// TIA Portal V20 export
DATA_BLOCK "DB020_Com LabView"   // DB20
{ S7_Optimized_Access := 'FALSE' }
// stored: AutoNumber false
   VAR
      E_Lebenszeichen : DInt := 0;   // E_Lebenszeichen
      E_Rückmeldung_Startfreigabe_Zwischenbefundung_erhalten : Bool;   // E_Rückmeldung_Startfreigabe_Zwischenbefundung_erhalten
      E_Rückmeldung_Zwischenbefundung_fertig : Bool;   // E_Rückmeldung_Zwischenbefundung_fertig
      "E_Messgerät ist bereit und verbunden" : Bool;   // E_Messgeräte_bereit
      "E_Messgerät ist Störungsfrei" : Bool;   // E_Messgerät ist Störungsfrei
      E_4_4 : Bool;
      E_4_5 : Bool;
      E_4_6 : Bool;
      E_4_7 : Bool;
      A_Lebenszeichen : DInt := 0;   // A_Lebenszeichen
      A_Startfreigabe_Zwischenbefundung : Bool;   // A_Startfreigabe_Zwischenbefundung
      A_Rückmeldung_Signal_Zwischenbfundung_erhalten : Bool;   // A_Rückmeldung_Signal_Zwischenbfundung_erhalten
      A_10_2 : Bool;
      A_10_3 : Bool;
      A_10_4 : Bool;
      A_10_5 : Bool;
      A_10_6 : Bool;
      A_10_7 : Bool;
      A_Betriebsart : Int := 0;   // Betriebsart Anlage 0=Aus , 1=Manuell, 2=Automatik, 3=Verwaltung, 4=Richten
      A_Steckzyklen_Soll : Int;   // A_Steckzyklen_Soll
      A_Steckzyklen_Ist : Int;   // A_Steckzyklen_Ist
      A_Achse_Istposition : Real := -0.96;   // A Achse Istposition in mm
      A_Achse_Drehmoment : Real := -0.96;   // A Achse Drehmoment in %
      A_Drehachse_Istposition : Real := -2.31;   // A Drehachse Istposition in °
      A_Drehachse_Drehmoment : Real := -2.31;   // A Drehachse Drehmoment in °
      A_Wegmessung_Ausgleichszylinder_Istwert : Real;   // A Wegmessung Ausgleichszylinder Istwert in mm
      A_Kraftsensor_Istwert : Real;   // A Kraftsensor Istwert in N
      A_Regelventil_Ausgleichszylinder_Istwert : Real;   // A Regelventil Ausgleichszylinder Istwert in mbar
      A_Regelventil_Überlastzylinder_Istwert : Real;   // A Regelventil Überlastzylinder Istwert in mbar
   END_VAR
BEGIN
END_DATA_BLOCK
